Fanuc KAREL source: kt00918.KL

-- PROVISIONAL review KL for V940-1; original PC SHA256 d24dd26e8268be05aa68e9185f413b3a059690dbebb20ce68373870985221c84
-- Incomplete behavior may be omitted. Consult companion uncertainty JSON. Do not deploy.
PROGRAM KT00918
%NOLOCKGROUP
VAR
  S1 : STRING[80]
  S2 : STRING[80]
  OUT : INTEGER
BEGIN
  -- V9_ZERO_TABLE_METADATA_HINT layout=0001; no indexed target words; source/name/runtime held
  -- UNRESOLVED_PC offsets 5-14; opcodes 3F,75
  -- UNRESOLVED_PC offsets 19-28; opcodes 3F,75
  -- UNRESOLVED_PC offsets 33-42; opcodes 3F,75
  -- UNRESOLVED_PC offsets 47-56; opcodes 3F,75
  -- UNRESOLVED_PC offsets 61-86; opcodes 27,22,2A,22,2A,76,23
  -- UNRESOLVED_PC offsets 91-95; opcodes 7F
END KT00918
